// Input block of T_RpcTarget.Add as sent over ADS.
TYPE ST_RpcAddParams :
STRUCT
  a : DINT;
  b : DINT;
END_STRUCT
END_TYPE

(* stored: Version 1.1.0.1, ProductVersion 3.1.4026.22
   DUT ST_RpcAddParams: Id {9fb974a3-0f95-43a7-a9a8-10bdaae70d91} *)
